RoboDK station: kukaiiwa_14.rdk

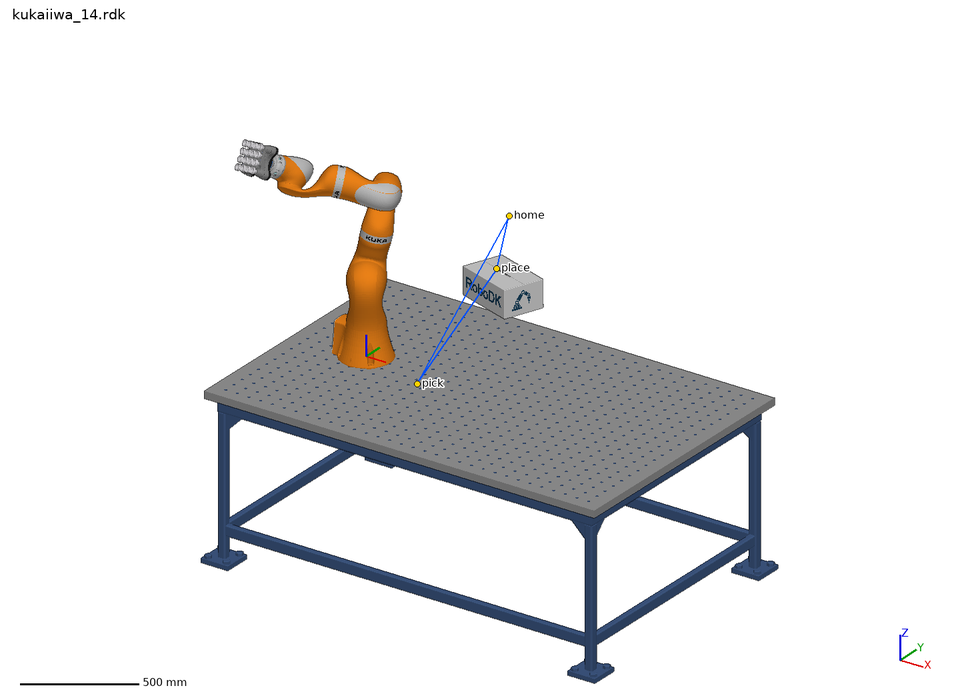
[picture v0: the station drawn from its stored meshes, robots at their saved joint values, targets as dots, program paths as lines]
Station kukaiiwa_14 (saved by RoboDK 6.0.6). Poses are relative to the parent item; angles as X-Y-Z fixed-axis rotations.
Station parameters (name, value as stored): LIN64
  - frame KUKA LBR iiwa 14 R820 Base at (0, 0, 0) mm
    - robot KUKA LBR iiwa 14 R820: 7 axes, payload 14 kg, reach 820 mm, repeatability 0.1 mm, weight 29.9 kg
        modified DH rows (alpha deg, a mm, theta deg, d mm): 0, 0, 0, 360; -90, 0, 0, 0; 90, 0, 0, 420; -90, 0, 0, 0; 90, 0, 0, 400; -90, 0, 0, 0; 90, 0, 0, 126
        joint limits [-170, -120, -170, -120, -170, -120, -175] to [170, 120, 170, 120, 170, 120, 175]; home [0, 0, 0, -90, 0, 0, 0]; saved at [32.597, 11.105, 0, -88.998, -53.999, 34.448, 80.368]
      - tool OnRobot VG10 Vacuum Gripper, TCP at (0, 0, 120.9) mm, size 145.4 x 145.4 x 118.3 mm
    - target home (Cartesian target) at (637.15, 135.96, 780) mm, rotated rx 0 ry 90 rz 0 deg; joints [19.207, 1.809, 0, -88.162, -89.914, 19.207, 89.909] of KUKA LBR iiwa 14 R820
    - target pick (Cartesian target) at (485.53, -320.08, 136.7) mm, rotated rx 172.18 ry 2.87 rz 96.39 deg; joints [-34.657, 41.315, 0, -96.09, 5.203, 34.923, 44.686] of KUKA LBR iiwa 14 R820
    - target place (Cartesian target) at (353.76, 451.22, 327.69) mm, rotated rx 172.99 ry 4.17 rz 166.28 deg; joints [52.309, 24.792, 0, -90.23, -1.123, 56.885, 66.322] of KUKA LBR iiwa 14 R820
  - object Table 2000x1200x800mm at (0, 0, 0) mm, size 2020 x 1340 x 800 mm, geometry from Table-2000x1200x800mm.sld
  - program Prog1 (10 instructions, listed below)
  - object Box 12x7in (Closed) at (501.61, 293.52, 196.73) mm, rotated rx -1.38 ry 0.66 rz 69.83 deg, size 199 x 305.1 x 133.7 mm, geometry from Box-12x7in-Closed.sld
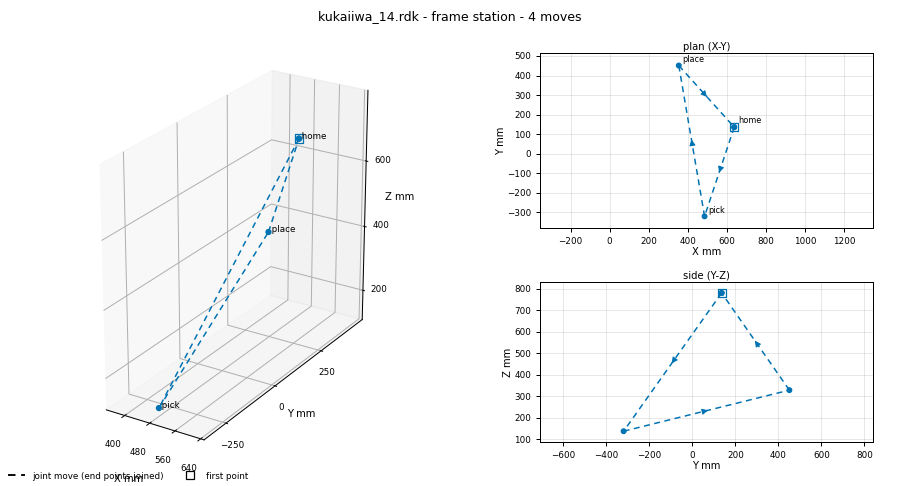
[picture p0: tool path of kukaiiwa_14.rdk in frame station, 4 of 4 moves have a stored position in this frame; points joined in program order, loops and branches not executed]

--- program Prog1 (robot KUKA LBR iiwa 14 R820) ---
  Set Ref.: KUKA LBR iiwa 14 R820 Base
  Set Tool: OnRobot VG10 Vacuum Gripper
  MoveJ (home)
  MoveJ (pick)
  Attach to OnRobot VG10 Vacuum Gripper
  MoveJ (place)
  Detach from OnRobot VG10 Vacuum Gripper
  MoveJ (home)
  Move Box 12x7in (Closed)
  Call Program1
